// TIA Portal V21 export
// export: Created 2026-11-10T19:11:37.5908756Z, ExportSetting WithDefaults, DisplayName Totally Integrated Automation Portal, DisplayVersion V21 Update 3, DisplayName STEP 7 Professional, DisplayVersion V21 Update 3, DisplayName STEP 7 Safety, DisplayVersion V21, DisplayName Tech WebApplication, DisplayVersion V21, DisplayName WinCC Basic/Comfort/Advanced, DisplayVersion V21 Update 3, DisplayName WinCC Unified, DisplayVersion V21 Update 3
DATA_BLOCK "DB_MCAT"   // DB24
// stored: AutoNumber true, DBAccessibleFromOPCUA true, DBAccessibleFromWebserver true, InstanceOfName MCAT, OfSystemLibElement MCAT, OfSystemLibVersion 2.1
"MCAT"
   // VAR_INPUT
   //    O_CMD : Bool;
   //    C_CMD : Bool;
   //    S_CMD : Bool;
   //    O_FB : Bool;
   //    C_FB : Bool;
   // END_VAR
   // VAR_OUTPUT
   //    OO : Bool;
   //    CO : Bool;
   //    OA : Bool;
   //    CA : Bool;
   //    Q : Bool;
   // END_VAR
   // VAR
   //    ET : DInt;
   //    PT : DInt;
   //    PREV_TIME : DWord;
   //    O_HIS : Bool;
   //    C_HIS : Bool;
   // END_VAR
BEGIN
END_DATA_BLOCK
